(* Logix 5000 project; controller _1407974_PSG_7315 vendor 1 type 14 code 154 rev 20.11; software revision 20.06; part 4 of 4 *)
(* tags used below, declared in another part *)
   AI_L_2_0_Pure_Steam_Conductivity : Analog_Input;
   AI_L_2_1_FW_Pressure : Analog_Input;
   AI_R_2_0_Pure_Steam_Temperature : Analog_Input;
   AI_R_2_1_Cond_Pure_Steam_Temperature : Analog_Input;
   Alarms_Warnings : AW;
   AO_R_4_0_Pure_Steam_Temperature : Analog_Output;
   AO_R_4_1_Available : Analog_Output;
   Cond_Pure_Steam_Conductivity_High : BOOL;
   Cond_Pure_Steam_Quality_OK_Latch : BOOL;
   Condensed_Pure_Steam_Warrnings_Disabled : Latched_Push_Button;
   Conductivity_Analzyer_Warmup_Delay_Timer : TIMER;
   DI_L_1_14_Feed_Water_Pump_Auto : ALIAS FOR DI_Local_1.14;
   DI_L_1_15_Feed_Water_Pump_Manual : ALIAS FOR DI_Local_1.15;
   DI_L_1_2_Pure_Steam_Analyzer_Fault : ALIAS FOR DI_Local_1.2;
   DI_Local_1 : INT;
   DI_Remote_1 : INT;
   DO_L_1_14_Feed_Water_Pump_Contactor : Discrete_Out;
   DO_L_1_15_Feed_Water_Pump_On_Light : Discrete_Out;
   DO_Local_1 : INT;
   DO_R_3_1_Primary_Level_Control_YV_4760 : Discrete_Out;
   DO_R_3_4_Degasser_Vent_YV_4255 : Discrete_Out;
   DO_R_3_5_FDW_TR : Discrete_Out;
   DO_Remote_3 : INT;
   F8_0_9 : REAL[10];
   Feed_Water_Pump_Delay_Timer : TIMER;
   Feedwater_Pressure_PID : PID;
   Lamp_Test : Push_Button;
   Local_Remote : Latched_Push_Button;
   Login_Popup : OIT_Popup;
   Login_Required_Popup : OIT_Popup;
   Maintenance_Mode : Latched_Push_Button;
   N7_0_9 : INT[10];
   Network_Ack_All : BOOL;
   Network_AI_L_2_0_Pure_Steam_Conductivity : REAL;
   Network_AI_L_2_1_Feedwater_Pressure : REAL;
   Network_AI_L_2_1_FW_Pressure_Scaled : DINT;
   Network_AI_R_2_0_Pure_Steam_Temperature : REAL;
   Network_AI_R_2_1_Cond_Pure_Steam_Temp : REAL;
   Network_AO_R_4_0_Pure_Steam_Man_Control : REAL;
   Network_AO_R_4_0_Pure_Steam_Temp_Control : REAL;
   Network_AO_R_4_1_Available_Manual : REAL;
   Network_AO_R_4_1_Available_Scaled : REAL;
   Network_Cond_PS_Temp_High_Set_Point : REAL;
   Network_DI_Local_1 : INT;
   Network_DI_Remote_1 : INT;
   Network_DO_Local_1 : INT;
   Network_DO_Remote_3 : INT;
   Network_Feedwater_Pressure_PID_KD : DINT;
   Network_Feedwater_Pressure_PID_KI : DINT;
   Network_Feedwater_Pressure_PID_KP : DINT;
   Network_Feedwater_Pressure_PID_SP : DINT;
   Network_FW_Low_Pressure_Warning_SP : DINT;
   Network_Input_Ack_All : BOOL;
   Network_Input_Silence : BOOL;
   Network_Input_Silence_ONS : BOOL;
   Network_Input_Start : BOOL;
   Network_Input_Start_ONS : BOOL;
   Network_Input_Stop : BOOL;
   Network_Input_Stop_ONS : BOOL;
   Network_PID_Ramp_Time_Seconds : DINT;
   Network_Pure_Steam_Conductivity_SetPoint : REAL;
   Network_Pure_Steam_Temp_High_Set_Point : REAL;
   Network_Pure_Steam_Temp_Lo_Set_Point : REAL;
   Network_Pure_Steam_Temp_PID_Gain : REAL;
   Network_Pure_Steam_Temp_PID_Rate : REAL;
   Network_Pure_Steam_Temp_PID_Reset : REAL;
   Network_Pure_Steam_Temperature_Set_Point : REAL;
   Network_Pure_Steam_Temporary_Set_Point : REAL;
   Network_Silence : BOOL;
   Network_Start : BOOL;
   Network_Status_Local_Remote : BOOL;
   Network_Status_Maintenance_Mode : BOOL;
   Network_Status_No_Active_Alarms : BOOL;
   Network_Status_No_Active_Warnings : BOOL;
   Network_Status_Unit_Cooling : BOOL;
   Network_Status_Unit_Filling : BOOL;
   Network_Status_Unit_Heating : BOOL;
   Network_Status_Unit_OFF : BOOL;
   Network_Status_Unit_ON : BOOL;
   Network_Status_Unit_Ready : BOOL;
   Network_Status_Unit_Running : BOOL;
   Network_Stop : BOOL;
   Netwrok_Input_Ack_All_ONS : BOOL;
   OIT : OIT_Connections;
   PID_Ramp_Time_Seconds : DINT;
   Pure_Steam_Temperature : PID;
   Read_PLC_Clock : DINT[7];
   Start_Stop_Popup : OIT_Popup;
   Unit_Status : Unit_Status;
   VFD_Relay_Input : BOOL;
   Warning_Cond_Pure_Steam_Analyzer_Fault : ALIAS FOR Alarms_Warnings.Latch_Bit[1].4;
   Warning_Cond_Pure_Steam_Analyzer_Timer : TIMER;
   Warning_Cond_Pure_Steam_Anlzr_Fault_Ack : ALIAS FOR Alarms_Warnings.Ack[1].4;
   Warning_Cond_Pure_Steam_Conduct_Timer : TIMER;
   Warning_Cond_Pure_Steam_Conductivity : ALIAS FOR Alarms_Warnings.Latch_Bit[1].3;
   Warning_Cond_Pure_Steam_Conductivity_Ack : ALIAS FOR Alarms_Warnings.Ack[1].3;
   Warning_Cond_Pure_Steam_Hi_Temp_Timer : TIMER;
   Warning_Cond_Pure_Steam_High_Temp : ALIAS FOR Alarms_Warnings.Latch_Bit[1].8;
   Warning_Cond_Pure_Steam_High_Temp_Ack : ALIAS FOR Alarms_Warnings.Ack[1].8;
   Warning_Feed_Water_Pump_Fault : ALIAS FOR Alarms_Warnings.Latch_Bit[1].1;
   Warning_Feed_Water_Pump_Fault_Ack : ALIAS FOR Alarms_Warnings.Ack[1].1;
   Warning_Feed_Water_Pump_Fault_Timer : TIMER;
(* MainProgram, continued *)

ROUTINE _100_Network_Buffer   (* ladder *)
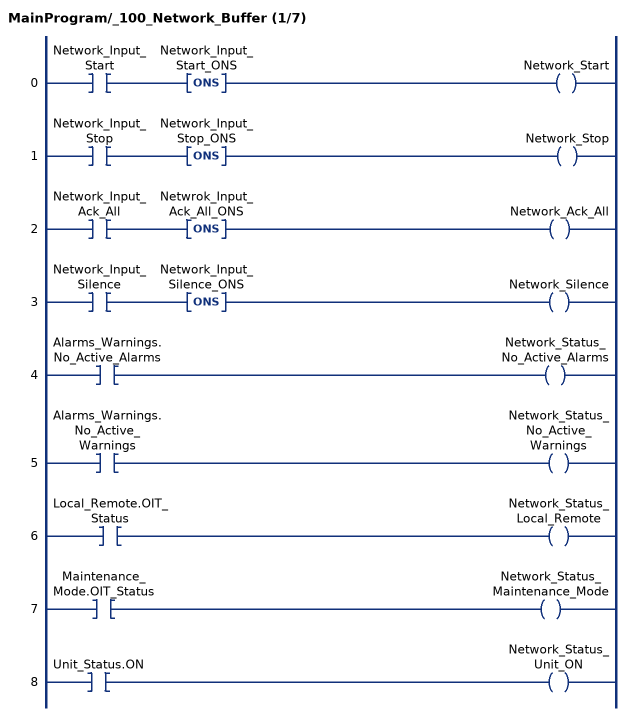
   0: XIC(Network_Input_Start)ONS(Network_Input_Start_ONS)OTE(Network_Start);
   1: XIC(Network_Input_Stop)ONS(Network_Input_Stop_ONS)OTE(Network_Stop);
   2: XIC(Network_Input_Ack_All)ONS(Netwrok_Input_Ack_All_ONS)OTE(Network_Ack_All);
   3: XIC(Network_Input_Silence)ONS(Network_Input_Silence_ONS)OTE(Network_Silence);
   4: XIC(Alarms_Warnings.No_Active_Alarms)OTE(Network_Status_No_Active_Alarms);
   5: XIC(Alarms_Warnings.No_Active_Warnings)OTE(Network_Status_No_Active_Warnings);
   6: XIC(Local_Remote.OIT_Status)OTE(Network_Status_Local_Remote);
   7: XIC(Maintenance_Mode.OIT_Status)OTE(Network_Status_Maintenance_Mode);
   8: XIC(Unit_Status.ON)OTE(Network_Status_Unit_ON);
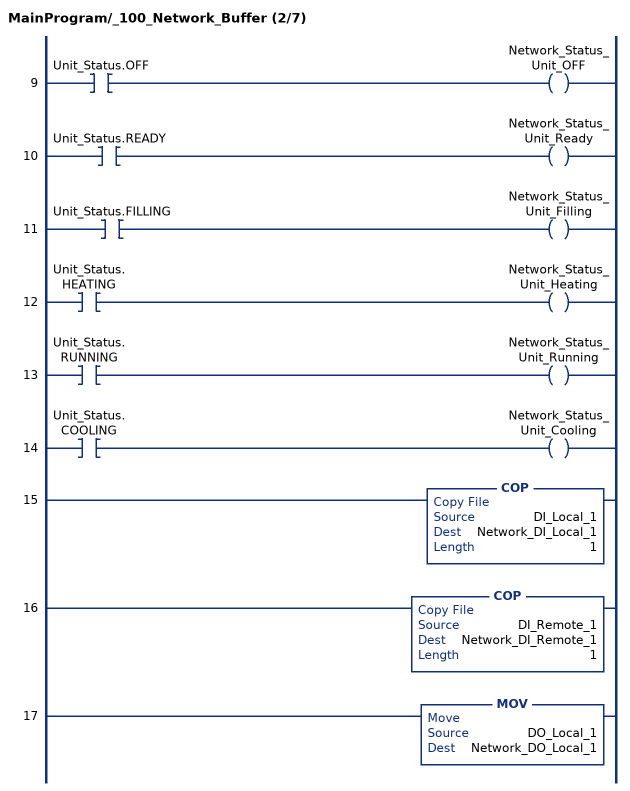
   9: XIC(Unit_Status.OFF)OTE(Network_Status_Unit_OFF);
   10: XIC(Unit_Status.READY)OTE(Network_Status_Unit_Ready);
   11: XIC(Unit_Status.FILLING)OTE(Network_Status_Unit_Filling);
   12: XIC(Unit_Status.HEATING)OTE(Network_Status_Unit_Heating);
   13: XIC(Unit_Status.RUNNING)OTE(Network_Status_Unit_Running);
   14: XIC(Unit_Status.COOLING)OTE(Network_Status_Unit_Cooling);
   15: COP(DI_Local_1,Network_DI_Local_1,1);
   16: COP(DI_Remote_1,Network_DI_Remote_1,1);
   17: MOV(DO_Local_1,Network_DO_Local_1);
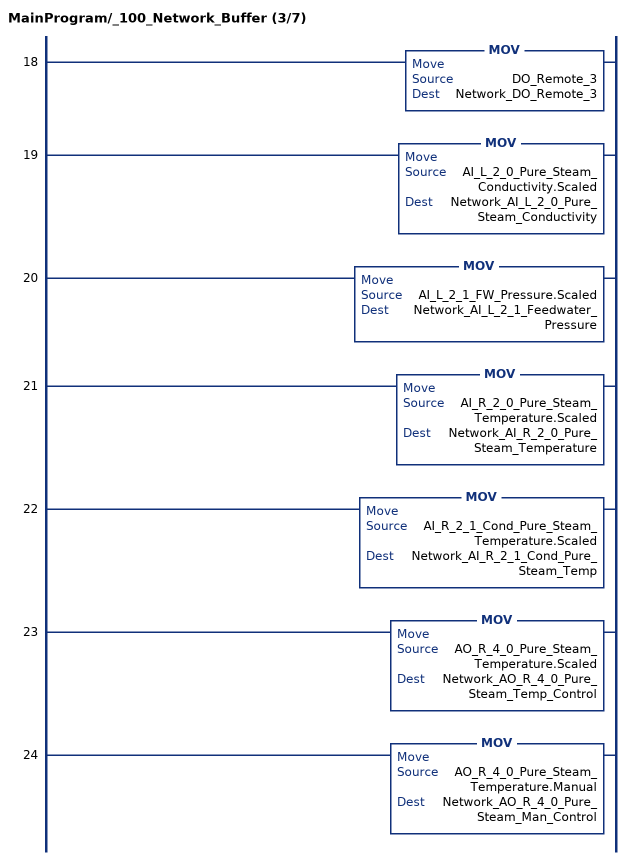
   18: MOV(DO_Remote_3,Network_DO_Remote_3);
   19: MOV(AI_L_2_0_Pure_Steam_Conductivity.Scaled,Network_AI_L_2_0_Pure_Steam_Conductivity);
   20: MOV(AI_L_2_1_FW_Pressure.Scaled,Network_AI_L_2_1_Feedwater_Pressure);
   21: MOV(AI_R_2_0_Pure_Steam_Temperature.Scaled,Network_AI_R_2_0_Pure_Steam_Temperature);
   22: MOV(AI_R_2_1_Cond_Pure_Steam_Temperature.Scaled,Network_AI_R_2_1_Cond_Pure_Steam_Temp);
   23: MOV(AO_R_4_0_Pure_Steam_Temperature.Scaled,Network_AO_R_4_0_Pure_Steam_Temp_Control);
   24: MOV(AO_R_4_0_Pure_Steam_Temperature.Manual,Network_AO_R_4_0_Pure_Steam_Man_Control);
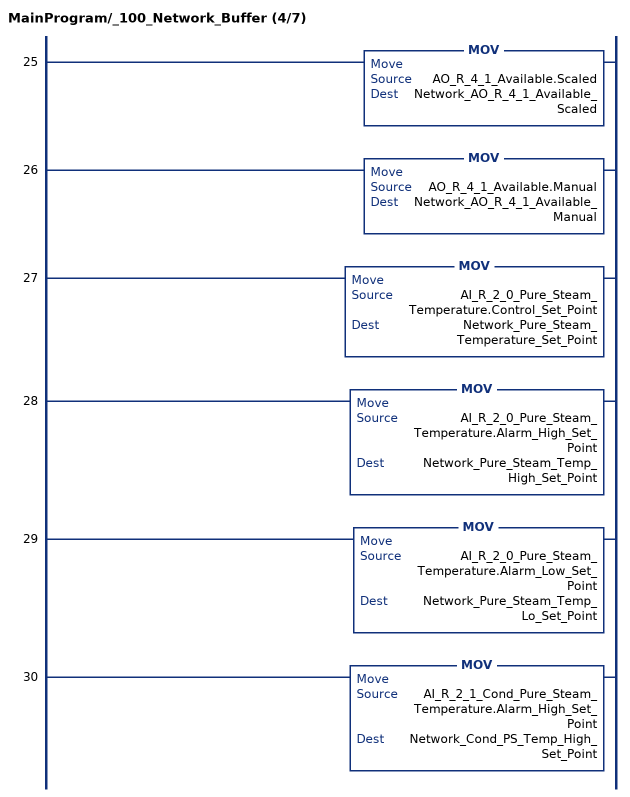
   25: MOV(AO_R_4_1_Available.Scaled,Network_AO_R_4_1_Available_Scaled);
   26: MOV(AO_R_4_1_Available.Manual,Network_AO_R_4_1_Available_Manual);
   27: MOV(AI_R_2_0_Pure_Steam_Temperature.Control_Set_Point,Network_Pure_Steam_Temperature_Set_Point);
   28: MOV(AI_R_2_0_Pure_Steam_Temperature.Alarm_High_Set_Point,Network_Pure_Steam_Temp_High_Set_Point);
   29: MOV(AI_R_2_0_Pure_Steam_Temperature.Alarm_Low_Set_Point,Network_Pure_Steam_Temp_Lo_Set_Point);
   30: MOV(AI_R_2_1_Cond_Pure_Steam_Temperature.Alarm_High_Set_Point,Network_Cond_PS_Temp_High_Set_Point);
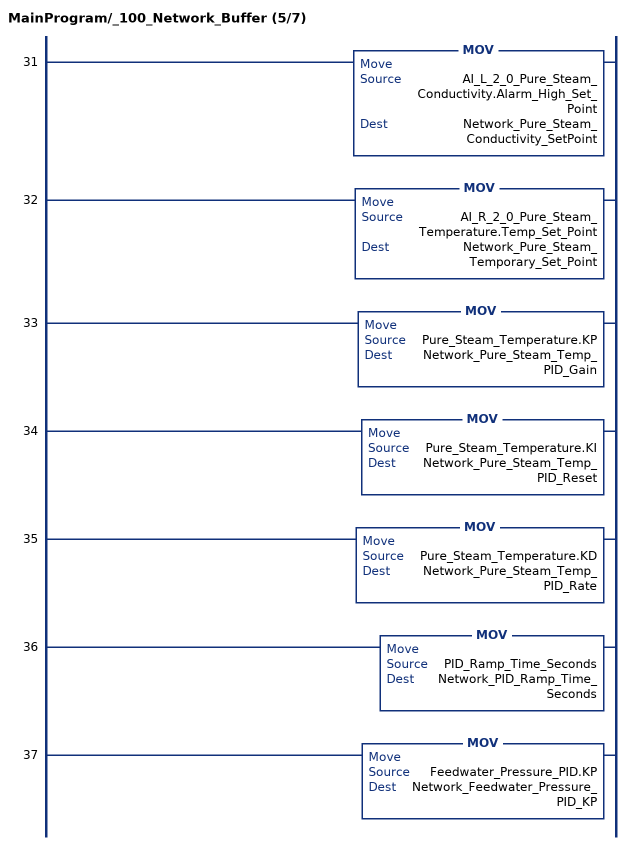
   31: MOV(AI_L_2_0_Pure_Steam_Conductivity.Alarm_High_Set_Point,Network_Pure_Steam_Conductivity_SetPoint);
   32: MOV(AI_R_2_0_Pure_Steam_Temperature.Temp_Set_Point,Network_Pure_Steam_Temporary_Set_Point);
   33: MOV(Pure_Steam_Temperature.KP,Network_Pure_Steam_Temp_PID_Gain);
   34: MOV(Pure_Steam_Temperature.KI,Network_Pure_Steam_Temp_PID_Reset);
   35: MOV(Pure_Steam_Temperature.KD,Network_Pure_Steam_Temp_PID_Rate);
   36: MOV(PID_Ramp_Time_Seconds,Network_PID_Ramp_Time_Seconds);
   37: MOV(Feedwater_Pressure_PID.KP,Network_Feedwater_Pressure_PID_KP);
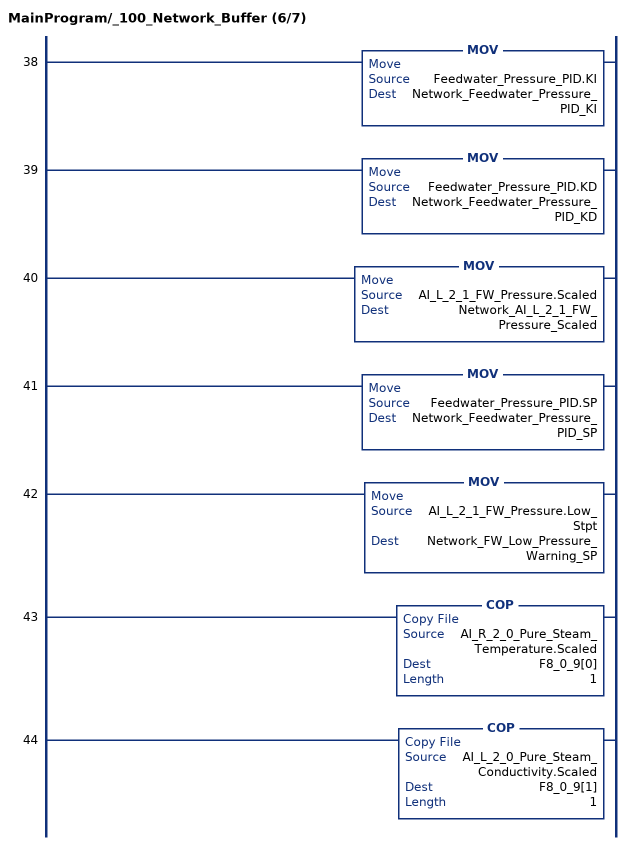
   38: MOV(Feedwater_Pressure_PID.KI,Network_Feedwater_Pressure_PID_KI);
   39: MOV(Feedwater_Pressure_PID.KD,Network_Feedwater_Pressure_PID_KD);
   40: MOV(AI_L_2_1_FW_Pressure.Scaled,Network_AI_L_2_1_FW_Pressure_Scaled);
   41: MOV(Feedwater_Pressure_PID.SP,Network_Feedwater_Pressure_PID_SP);
   42: MOV(AI_L_2_1_FW_Pressure.Low_Stpt,Network_FW_Low_Pressure_Warning_SP);
   43: COP(AI_R_2_0_Pure_Steam_Temperature.Scaled,F8_0_9[0],1);
   44: COP(AI_L_2_0_Pure_Steam_Conductivity.Scaled,F8_0_9[1],1);
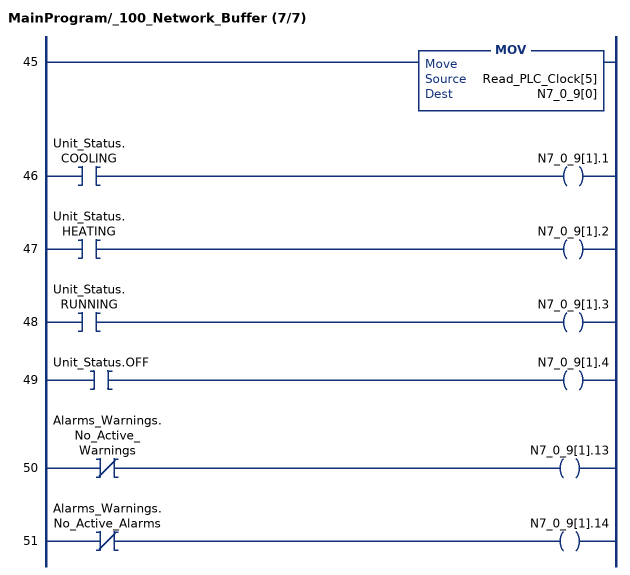
   45: MOV(Read_PLC_Clock[5],N7_0_9[0]);
   46: XIC(Unit_Status.COOLING)OTE(N7_0_9[1].1);
   47: XIC(Unit_Status.HEATING)OTE(N7_0_9[1].2);
   48: XIC(Unit_Status.RUNNING)OTE(N7_0_9[1].3);
   49: XIC(Unit_Status.OFF)OTE(N7_0_9[1].4);
   50: XIO(Alarms_Warnings.No_Active_Warnings)OTE(N7_0_9[1].13);
   51: XIO(Alarms_Warnings.No_Active_Alarms)OTE(N7_0_9[1].14);
END_ROUTINE

ROUTINE _110_Calls   (* ladder *)
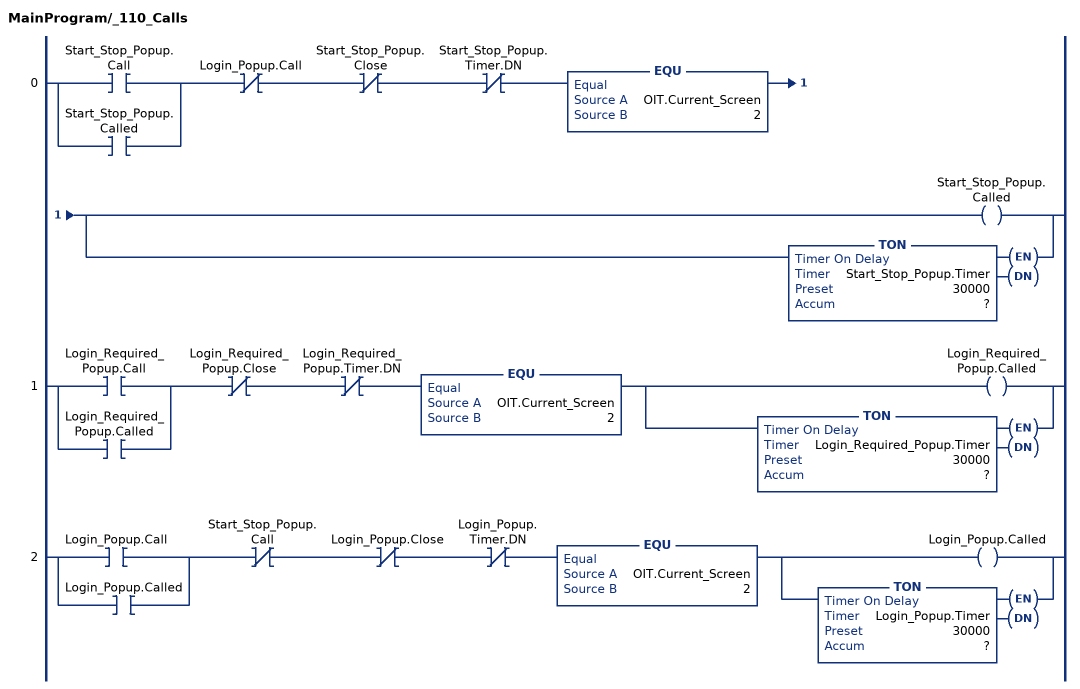
   0: [XIC(Start_Stop_Popup.Call) ,XIC(Start_Stop_Popup.Called) ]XIO(Login_Popup.Call)XIO(Start_Stop_Popup.Close)XIO(Start_Stop_Popup.Timer.DN)EQU(OIT.Current_Screen,2)[OTE(Start_Stop_Popup.Called) ,TON(Start_Stop_Popup.Timer,?,?) ];
   1: [XIC(Login_Required_Popup.Call) ,XIC(Login_Required_Popup.Called) ]XIO(Login_Required_Popup.Close)XIO(Login_Required_Popup.Timer.DN)EQU(OIT.Current_Screen,2)[OTE(Login_Required_Popup.Called) ,TON(Login_Required_Popup.Timer,?,?) ];
   2: [XIC(Login_Popup.Call) ,XIC(Login_Popup.Called) ]XIO(Start_Stop_Popup.Call)XIO(Login_Popup.Close)XIO(Login_Popup.Timer.DN)EQU(OIT.Current_Screen,2)[OTE(Login_Popup.Called) ,TON(Login_Popup.Timer,?,?) ];
END_ROUTINE

ROUTINE _120_Option_Condensed_Pure_Steam   (* ladder *)
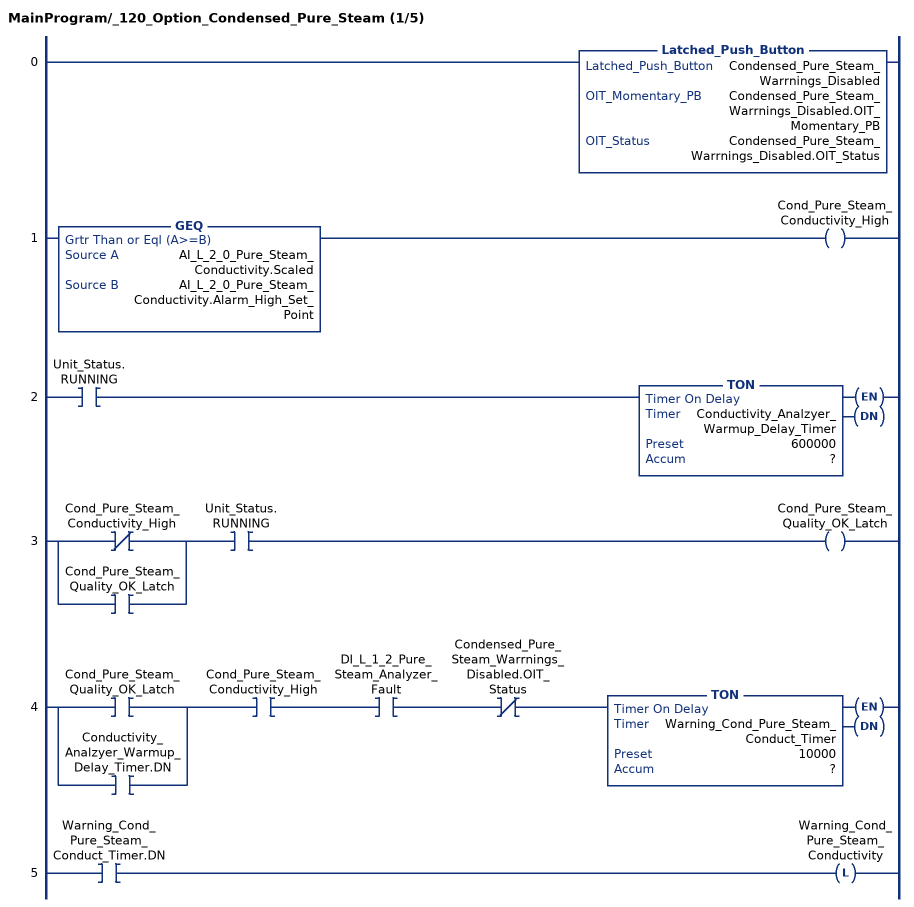
   0: Latched_Push_Button(Condensed_Pure_Steam_Warrnings_Disabled,Condensed_Pure_Steam_Warrnings_Disabled.OIT_Momentary_PB,Condensed_Pure_Steam_Warrnings_Disabled.OIT_Status);
   1: GEQ(AI_L_2_0_Pure_Steam_Conductivity.Scaled,AI_L_2_0_Pure_Steam_Conductivity.Alarm_High_Set_Point)OTE(Cond_Pure_Steam_Conductivity_High);
   2: XIC(Unit_Status.RUNNING)TON(Conductivity_Analzyer_Warmup_Delay_Timer,?,?);
   3: [XIO(Cond_Pure_Steam_Conductivity_High) ,XIC(Cond_Pure_Steam_Quality_OK_Latch) ]XIC(Unit_Status.RUNNING)OTE(Cond_Pure_Steam_Quality_OK_Latch);
   4: [XIC(Cond_Pure_Steam_Quality_OK_Latch) ,XIC(Conductivity_Analzyer_Warmup_Delay_Timer.DN) ]XIC(Cond_Pure_Steam_Conductivity_High)XIC(DI_L_1_2_Pure_Steam_Analyzer_Fault)XIO(Condensed_Pure_Steam_Warrnings_Disabled.OIT_Status)TON(Warning_Cond_Pure_Steam_Conduct_Timer,?,?);
   5: XIC(Warning_Cond_Pure_Steam_Conduct_Timer.DN)OTL(Warning_Cond_Pure_Steam_Conductivity);
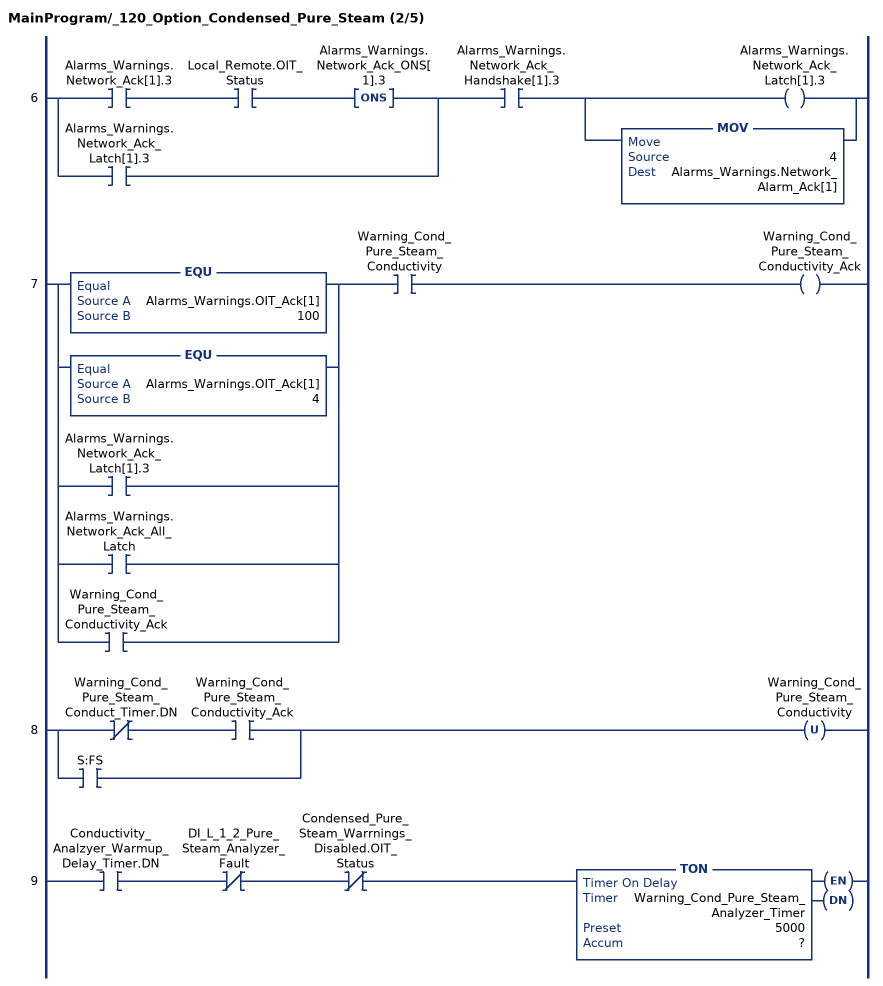
   6: [XIC(Alarms_Warnings.Network_Ack[1].3) XIC(Local_Remote.OIT_Status) ONS(Alarms_Warnings.Network_Ack_ONS[1].3) ,XIC(Alarms_Warnings.Network_Ack_Latch[1].3) ]XIC(Alarms_Warnings.Network_Ack_Handshake[1].3)[OTE(Alarms_Warnings.Network_Ack_Latch[1].3) ,MOV(4,Alarms_Warnings.Network_Alarm_Ack[1]) ];
   7: [EQU(Alarms_Warnings.OIT_Ack[1],100) ,EQU(Alarms_Warnings.OIT_Ack[1],4) ,XIC(Alarms_Warnings.Network_Ack_Latch[1].3) ,XIC(Alarms_Warnings.Network_Ack_All_Latch) ,XIC(Warning_Cond_Pure_Steam_Conductivity_Ack) ]XIC(Warning_Cond_Pure_Steam_Conductivity)OTE(Warning_Cond_Pure_Steam_Conductivity_Ack);
   8: [XIO(Warning_Cond_Pure_Steam_Conduct_Timer.DN) XIC(Warning_Cond_Pure_Steam_Conductivity_Ack) ,XIC(S:FS) ]OTU(Warning_Cond_Pure_Steam_Conductivity);
   9: XIC(Conductivity_Analzyer_Warmup_Delay_Timer.DN)XIO(DI_L_1_2_Pure_Steam_Analyzer_Fault)XIO(Condensed_Pure_Steam_Warrnings_Disabled.OIT_Status)TON(Warning_Cond_Pure_Steam_Analyzer_Timer,?,?);
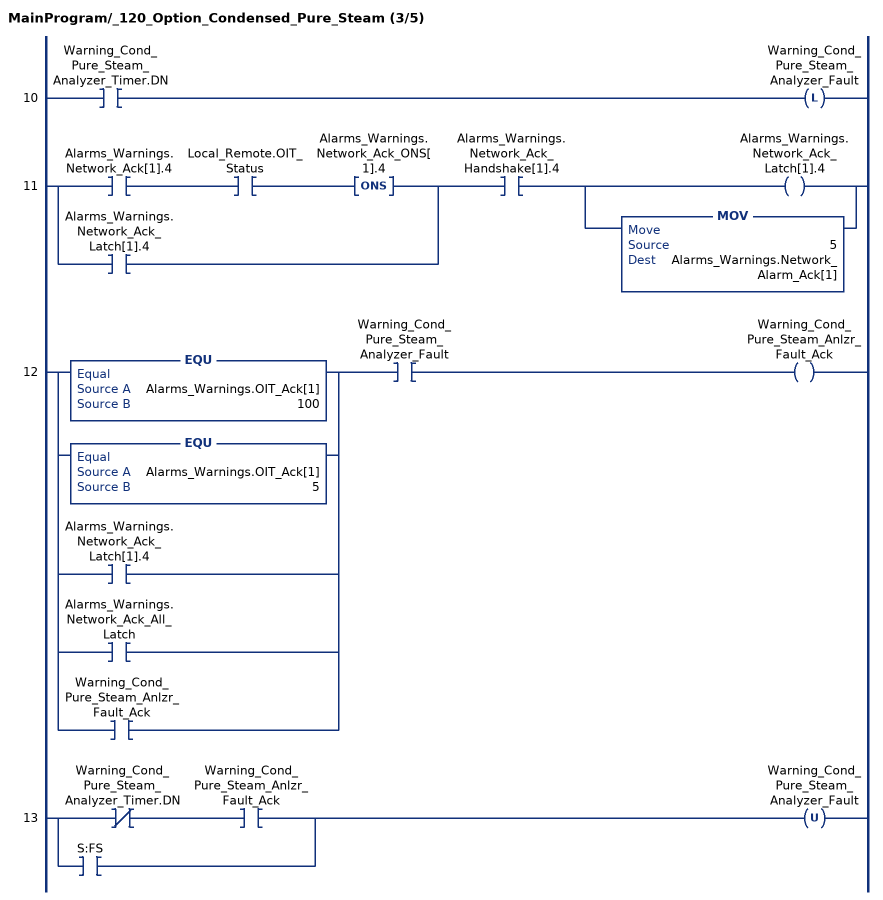
   10: XIC(Warning_Cond_Pure_Steam_Analyzer_Timer.DN)OTL(Warning_Cond_Pure_Steam_Analyzer_Fault);
   11: [XIC(Alarms_Warnings.Network_Ack[1].4) XIC(Local_Remote.OIT_Status) ONS(Alarms_Warnings.Network_Ack_ONS[1].4) ,XIC(Alarms_Warnings.Network_Ack_Latch[1].4) ]XIC(Alarms_Warnings.Network_Ack_Handshake[1].4)[OTE(Alarms_Warnings.Network_Ack_Latch[1].4) ,MOV(5,Alarms_Warnings.Network_Alarm_Ack[1]) ];
   12: [EQU(Alarms_Warnings.OIT_Ack[1],100) ,EQU(Alarms_Warnings.OIT_Ack[1],5) ,XIC(Alarms_Warnings.Network_Ack_Latch[1].4) ,XIC(Alarms_Warnings.Network_Ack_All_Latch) ,XIC(Warning_Cond_Pure_Steam_Anlzr_Fault_Ack) ]XIC(Warning_Cond_Pure_Steam_Analyzer_Fault)OTE(Warning_Cond_Pure_Steam_Anlzr_Fault_Ack);
   13: [XIO(Warning_Cond_Pure_Steam_Analyzer_Timer.DN) XIC(Warning_Cond_Pure_Steam_Anlzr_Fault_Ack) ,XIC(S:FS) ]OTU(Warning_Cond_Pure_Steam_Analyzer_Fault);
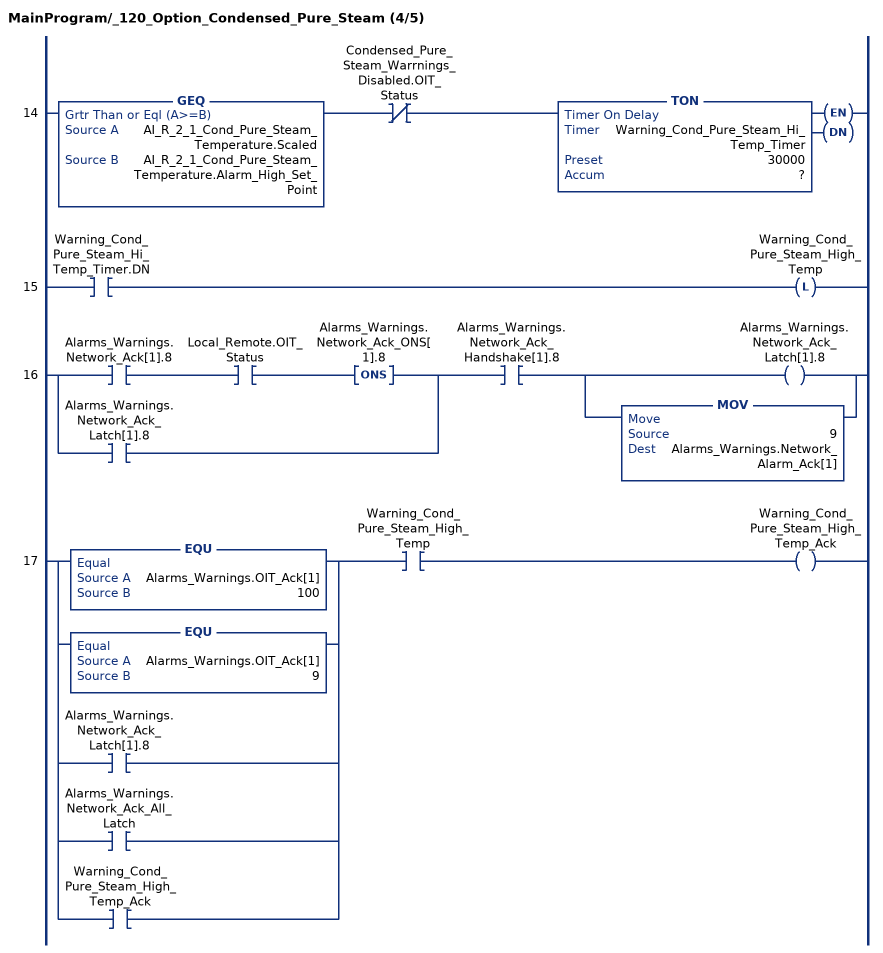
   14: GEQ(AI_R_2_1_Cond_Pure_Steam_Temperature.Scaled,AI_R_2_1_Cond_Pure_Steam_Temperature.Alarm_High_Set_Point)XIO(Condensed_Pure_Steam_Warrnings_Disabled.OIT_Status)TON(Warning_Cond_Pure_Steam_Hi_Temp_Timer,?,?);
   15: XIC(Warning_Cond_Pure_Steam_Hi_Temp_Timer.DN)OTL(Warning_Cond_Pure_Steam_High_Temp);
   16: [XIC(Alarms_Warnings.Network_Ack[1].8) XIC(Local_Remote.OIT_Status) ONS(Alarms_Warnings.Network_Ack_ONS[1].8) ,XIC(Alarms_Warnings.Network_Ack_Latch[1].8) ]XIC(Alarms_Warnings.Network_Ack_Handshake[1].8)[OTE(Alarms_Warnings.Network_Ack_Latch[1].8) ,MOV(9,Alarms_Warnings.Network_Alarm_Ack[1]) ];
   17: [EQU(Alarms_Warnings.OIT_Ack[1],100) ,EQU(Alarms_Warnings.OIT_Ack[1],9) ,XIC(Alarms_Warnings.Network_Ack_Latch[1].8) ,XIC(Alarms_Warnings.Network_Ack_All_Latch) ,XIC(Warning_Cond_Pure_Steam_High_Temp_Ack) ]XIC(Warning_Cond_Pure_Steam_High_Temp)OTE(Warning_Cond_Pure_Steam_High_Temp_Ack);
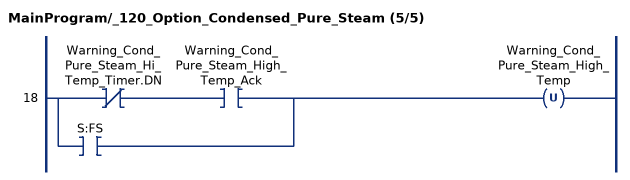
   18: [XIO(Warning_Cond_Pure_Steam_Hi_Temp_Timer.DN) XIC(Warning_Cond_Pure_Steam_High_Temp_Ack) ,XIC(S:FS) ]OTU(Warning_Cond_Pure_Steam_High_Temp);
END_ROUTINE

ROUTINE _130_Option_Feed_Water_Pump   (* ladder *)
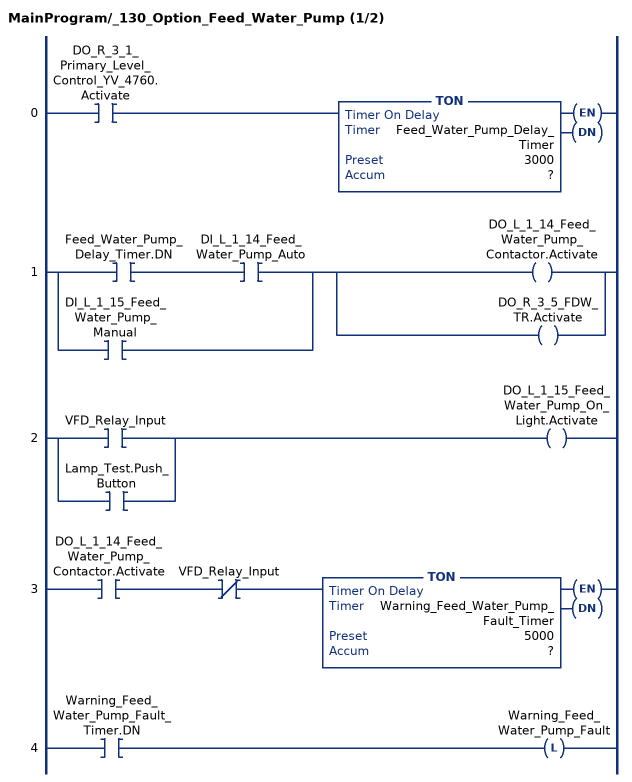
   0: XIC(DO_R_3_1_Primary_Level_Control_YV_4760.Activate)TON(Feed_Water_Pump_Delay_Timer,?,?);
   1: [XIC(Feed_Water_Pump_Delay_Timer.DN) XIC(DI_L_1_14_Feed_Water_Pump_Auto) ,XIC(DI_L_1_15_Feed_Water_Pump_Manual) ][OTE(DO_L_1_14_Feed_Water_Pump_Contactor.Activate) ,OTE(DO_R_3_5_FDW_TR.Activate) ];
   2: [XIC(VFD_Relay_Input) ,XIC(Lamp_Test.Push_Button) ]OTE(DO_L_1_15_Feed_Water_Pump_On_Light.Activate);
   3: XIC(DO_L_1_14_Feed_Water_Pump_Contactor.Activate)XIO(VFD_Relay_Input)TON(Warning_Feed_Water_Pump_Fault_Timer,?,?);
   4: XIC(Warning_Feed_Water_Pump_Fault_Timer.DN)OTL(Warning_Feed_Water_Pump_Fault);
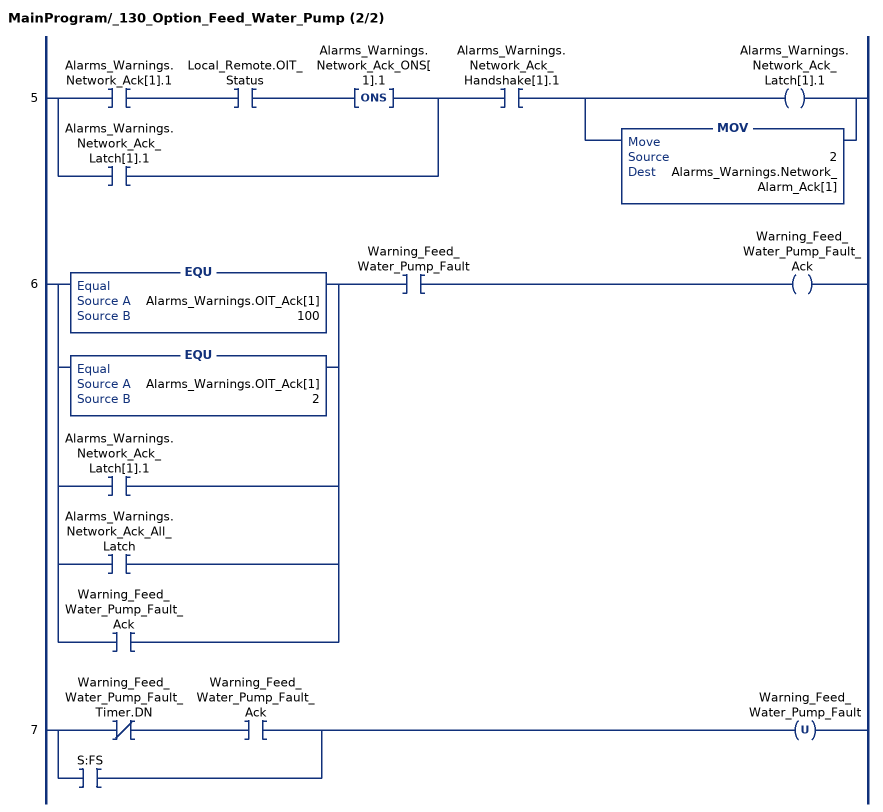
   5: [XIC(Alarms_Warnings.Network_Ack[1].1) XIC(Local_Remote.OIT_Status) ONS(Alarms_Warnings.Network_Ack_ONS[1].1) ,XIC(Alarms_Warnings.Network_Ack_Latch[1].1) ]XIC(Alarms_Warnings.Network_Ack_Handshake[1].1)[OTE(Alarms_Warnings.Network_Ack_Latch[1].1) ,MOV(2,Alarms_Warnings.Network_Alarm_Ack[1]) ];
   6: [EQU(Alarms_Warnings.OIT_Ack[1],100) ,EQU(Alarms_Warnings.OIT_Ack[1],2) ,XIC(Alarms_Warnings.Network_Ack_Latch[1].1) ,XIC(Alarms_Warnings.Network_Ack_All_Latch) ,XIC(Warning_Feed_Water_Pump_Fault_Ack) ]XIC(Warning_Feed_Water_Pump_Fault)OTE(Warning_Feed_Water_Pump_Fault_Ack);
   7: [XIO(Warning_Feed_Water_Pump_Fault_Timer.DN) XIC(Warning_Feed_Water_Pump_Fault_Ack) ,XIC(S:FS) ]OTU(Warning_Feed_Water_Pump_Fault);
END_ROUTINE

ROUTINE _140_Option_Feed_Water_Degasser   (* ladder *)
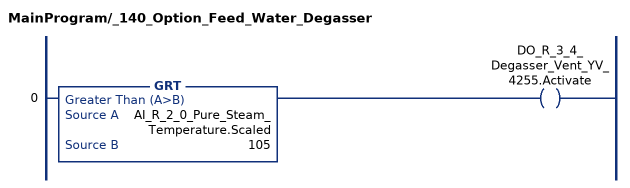
   0: GRT(AI_R_2_0_Pure_Steam_Temperature.Scaled,105)OTE(DO_R_3_4_Degasser_Vent_YV_4255.Activate);
END_ROUTINE
END_PROGRAM
